(* IEC 61131-3 sources: ZPLC/packages/zplc-ide/plant-scenes/colour-separation, 2 files *)

(* ---- reference.st ---- *)
PROGRAM ColourSeparation
VAR_INPUT
    Start     AT %I0.0 : BOOL;
    Waiting   AT %I0.1 : BOOL;
    IsRed     AT %I0.2 : BOOL;
    Extended  AT %I0.3 : BOOL;
    Retracted AT %I0.4 : BOOL;
END_VAR
VAR_OUTPUT
    RunIn     AT %Q0.0 : BOOL;
    RunOut    AT %Q0.1 : BOOL;
    RunSide   AT %Q0.2 : BOOL;
    Hold      AT %Q0.3 : BOOL;
    Push      AT %Q0.4 : BOOL;
    Busy      AT %Q0.5 : BOOL;
    Done      AT %Q0.6 : BOOL;
END_VAR
VAR
    Active  : BOOL;
    State   : INT;
    Red     : BOOL;
    Handled : INT;
    Settle  : TON;
    Clear   : TON;
END_VAR

IF Start THEN
    Active := TRUE;
END_IF;

(* the workpiece must lie still against the blade before its colour is read; after the
   release it must have left the blade before the blade holds again *)
Settle(IN := Waiting AND State = 0, PT := T#300ms);
Clear(IN := State = 3 AND NOT Waiting, PT := T#1500ms);

(* one state per step: 0 wait for a workpiece, 1 push it out, 2 pull the plate back,
   3 let a blue one go by *)
CASE State OF
    0:
        IF Active AND Settle.Q THEN
            Red := IsRed;
            IF Red THEN
                State := 1;
            ELSE
                State := 3;
            END_IF;
        END_IF;
    1:
        IF Extended THEN
            State := 2;
        END_IF;
    2:
        IF Retracted THEN
            Handled := Handled + 1;
            State := 0;
        END_IF;
    3:
        IF Clear.Q THEN
            Handled := Handled + 1;
            State := 0;
        END_IF;
END_CASE;

RunIn   := Active;
RunOut  := Active;
RunSide := Active;
(* the blade lets a blue workpiece go and holds everything else *)
Hold    := Active AND State <> 3;
Push    := State = 1;
Done    := Handled >= 8;
Busy    := Active AND NOT Done;

END_PROGRAM

(* ---- starter.st ---- *)
PROGRAM ColourSeparation
VAR_INPUT
    Start     AT %I0.0 : BOOL;  (* StartButton.pressed: start the line *)
    Waiting   AT %I0.1 : BOOL;  (* EyeStop.detect: a workpiece waits at the stop blade *)
    IsRed     AT %I0.2 : BOOL;  (* Colour1.match: the workpiece in the beam is red *)
    Extended  AT %I0.3 : BOOL;  (* Pusher1.extended: the plate is fully out *)
    Retracted AT %I0.4 : BOOL;  (* Pusher1.retracted: the plate is fully back *)
END_VAR
VAR_OUTPUT
    RunIn     AT %Q0.0 : BOOL;  (* Infeed.run: run the infeed belt *)
    RunOut    AT %Q0.1 : BOOL;  (* Outfeed.run: run the belt that ends in BlueBin *)
    RunSide   AT %Q0.2 : BOOL;  (* SideBelt.run: run the belt that ends in RedBin *)
    Hold      AT %Q0.3 : BOOL;  (* Stop1.extend: the blade holds a workpiece while true *)
    Push      AT %Q0.4 : BOOL;  (* Pusher1.extend: push sideways while true, retract when false *)
    Busy      AT %Q0.5 : BOOL;  (* Beacon.amber: the line is running *)
    Done      AT %Q0.6 : BOOL;  (* Beacon.green: lit when eight workpieces are sorted *)
END_VAR

(* Goal: a press of the start button runs the three belts. Eight workpieces,
   red or blue, arrive one at a time on the infeed. The blade stops each one
   in front of the colour sensor. Wait until it lies still, then read IsRed.
   A red one is pushed onto the side belt: extend the pusher until Extended,
   then retract it and wait for Retracted. A blue one is released by the blade
   and rides on to the outfeed. Hold the blade again once the workpiece has
   gone. Light Busy while the line runs and Done after the eighth workpiece. *)

END_PROGRAM
